// TIA Portal V20 export
// export: Created 2026-10-20T12:51:39.2775664Z, ExportSetting WithDefaults, DisplayName Totally Integrated Automation Portal, DisplayVersion V20 Update 6, DisplayName TIA Portal Openness, DisplayVersion V20 Update 6, DisplayName TIA Portal Version Control Interface, DisplayVersion V20 Update 6, DisplayName SINAMICS Startdrive Advanced, DisplayVersion V20 SP1, DisplayName SINAMICS Startdrive G130, G150, S120, S150, SINAMICS MV, G220, S200, S210, DisplayVersion V20 SP1, DisplayName SINAMICS Startdrive G110M, G120, G120C, G120D, G120P, G115D, DisplayVersion V20 SP1, DisplayName STEP 7 Professional, DisplayVersion V20 Update 6, DisplayName STEP 7 Safety, DisplayVersion V20 Update 2, DisplayName WinCC Basic/Comfort/Advanced, DisplayVersion V20 Update 6, DisplayName WinCC Unified, DisplayVersion V20 Update 6
FUNCTION "Bypass assignments_2" : Void   // FC36, F_LAD
{ S7_Optimized_Access := 'TRUE' }
VERSION : 0.1
// stored: AutoNumber true, IsIECCheckEnabled false, UDAEnableTagReadback false
BEGIN

REGION Network 1
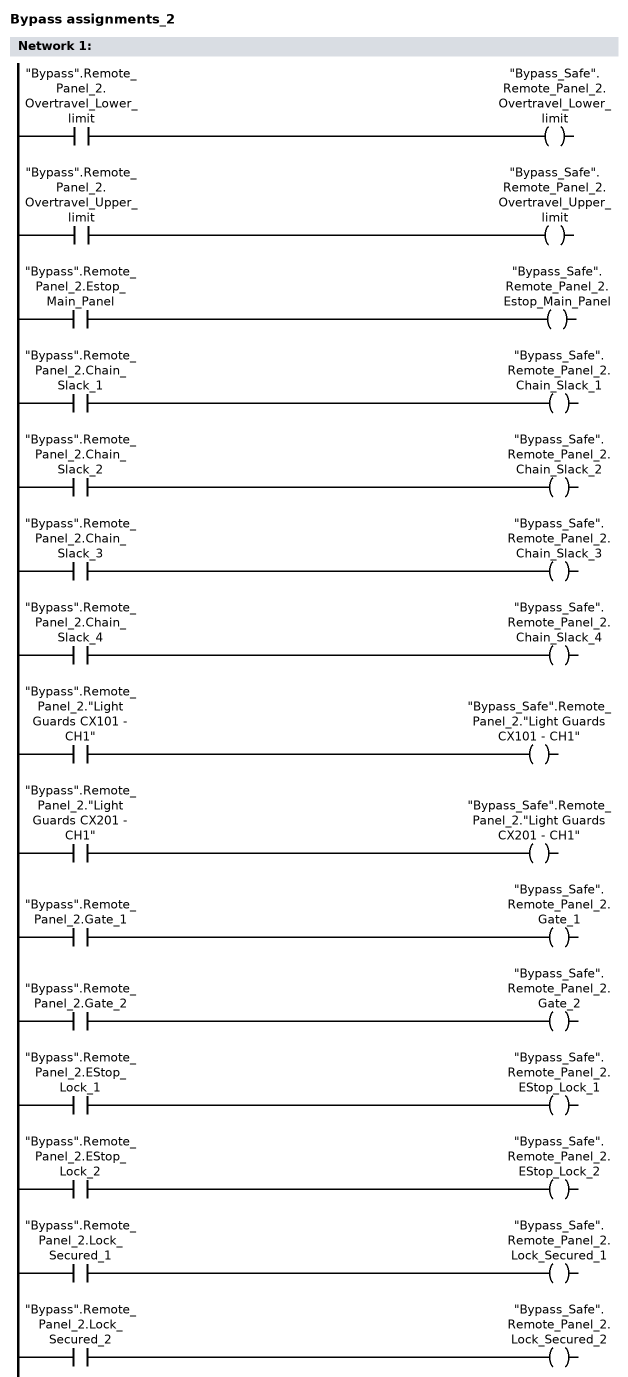
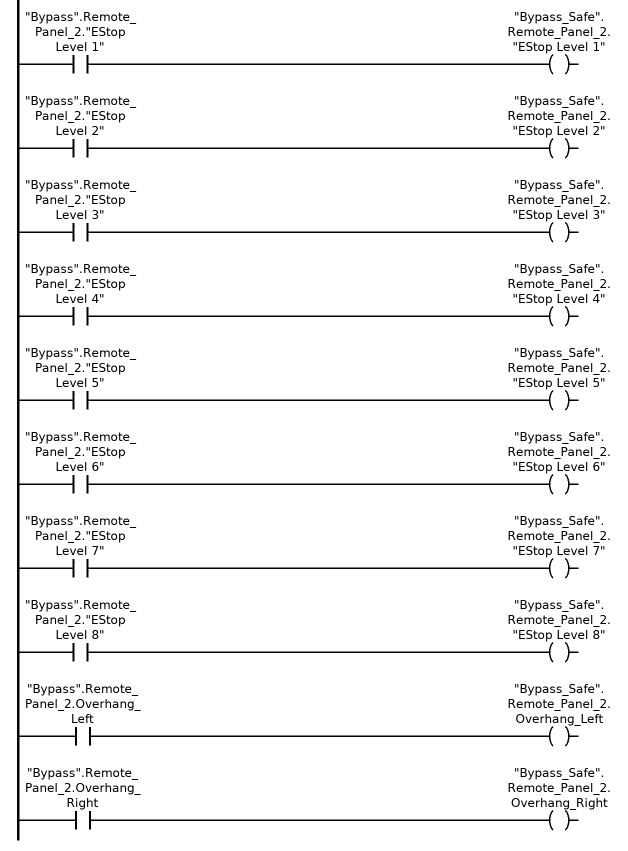
   RUNG wire#powerrail
      Contact( "Bypass".Remote_Panel_2.Overtravel_Lower_limit )
      Coil( "Bypass_Safe".Remote_Panel_2.Overtravel_Lower_limit )
   END_RUNG
   RUNG wire#powerrail
      Contact( "Bypass".Remote_Panel_2.Overtravel_Upper_limit )
      Coil( "Bypass_Safe".Remote_Panel_2.Overtravel_Upper_limit )
   END_RUNG
   RUNG wire#powerrail
      Contact( "Bypass".Remote_Panel_2.Estop_Main_Panel )
      Coil( "Bypass_Safe".Remote_Panel_2.Estop_Main_Panel )
   END_RUNG
   RUNG wire#powerrail
      Contact( "Bypass".Remote_Panel_2.Chain_Slack_1 )
      Coil( "Bypass_Safe".Remote_Panel_2.Chain_Slack_1 )
   END_RUNG
   RUNG wire#powerrail
      Contact( "Bypass".Remote_Panel_2.Chain_Slack_2 )
      Coil( "Bypass_Safe".Remote_Panel_2.Chain_Slack_2 )
   END_RUNG
   RUNG wire#powerrail
      Contact( "Bypass".Remote_Panel_2.Chain_Slack_3 )
      Coil( "Bypass_Safe".Remote_Panel_2.Chain_Slack_3 )
   END_RUNG
   RUNG wire#powerrail
      Contact( "Bypass".Remote_Panel_2.Chain_Slack_4 )
      Coil( "Bypass_Safe".Remote_Panel_2.Chain_Slack_4 )
   END_RUNG
   RUNG wire#powerrail
      Contact( "Bypass".Remote_Panel_2."Light Guards CX101 - CH1" )
      Coil( "Bypass_Safe".Remote_Panel_2."Light Guards CX101 - CH1" )
   END_RUNG
   RUNG wire#powerrail
      Contact( "Bypass".Remote_Panel_2."Light Guards CX201 - CH1" )
      Coil( "Bypass_Safe".Remote_Panel_2."Light Guards CX201 - CH1" )
   END_RUNG
   RUNG wire#powerrail
      Contact( "Bypass".Remote_Panel_2.Gate_1 )
      Coil( "Bypass_Safe".Remote_Panel_2.Gate_1 )
   END_RUNG
   RUNG wire#powerrail
      Contact( "Bypass".Remote_Panel_2.Gate_2 )
      Coil( "Bypass_Safe".Remote_Panel_2.Gate_2 )
   END_RUNG
   RUNG wire#powerrail
      Contact( "Bypass".Remote_Panel_2.EStop_Lock_1 )
      Coil( "Bypass_Safe".Remote_Panel_2.EStop_Lock_1 )
   END_RUNG
   RUNG wire#powerrail
      Contact( "Bypass".Remote_Panel_2.EStop_Lock_2 )
      Coil( "Bypass_Safe".Remote_Panel_2.EStop_Lock_2 )
   END_RUNG
   RUNG wire#powerrail
      Contact( "Bypass".Remote_Panel_2.Lock_Secured_1 )
      Coil( "Bypass_Safe".Remote_Panel_2.Lock_Secured_1 )
   END_RUNG
   RUNG wire#powerrail
      Contact( "Bypass".Remote_Panel_2.Lock_Secured_2 )
      Coil( "Bypass_Safe".Remote_Panel_2.Lock_Secured_2 )
   END_RUNG
   RUNG wire#powerrail
      Contact( "Bypass".Remote_Panel_2."EStop Level 1" )
      Coil( "Bypass_Safe".Remote_Panel_2."EStop Level 1" )
   END_RUNG
   RUNG wire#powerrail
      Contact( "Bypass".Remote_Panel_2."EStop Level 2" )
      Coil( "Bypass_Safe".Remote_Panel_2."EStop Level 2" )
   END_RUNG
   RUNG wire#powerrail
      Contact( "Bypass".Remote_Panel_2."EStop Level 3" )
      Coil( "Bypass_Safe".Remote_Panel_2."EStop Level 3" )
   END_RUNG
   RUNG wire#powerrail
      Contact( "Bypass".Remote_Panel_2."EStop Level 4" )
      Coil( "Bypass_Safe".Remote_Panel_2."EStop Level 4" )
   END_RUNG
   RUNG wire#powerrail
      Contact( "Bypass".Remote_Panel_2."EStop Level 5" )
      Coil( "Bypass_Safe".Remote_Panel_2."EStop Level 5" )
   END_RUNG
   RUNG wire#powerrail
      Contact( "Bypass".Remote_Panel_2."EStop Level 6" )
      Coil( "Bypass_Safe".Remote_Panel_2."EStop Level 6" )
   END_RUNG
   RUNG wire#powerrail
      Contact( "Bypass".Remote_Panel_2."EStop Level 7" )
      Coil( "Bypass_Safe".Remote_Panel_2."EStop Level 7" )
   END_RUNG
   RUNG wire#powerrail
      Contact( "Bypass".Remote_Panel_2."EStop Level 8" )
      Coil( "Bypass_Safe".Remote_Panel_2."EStop Level 8" )
   END_RUNG
   RUNG wire#powerrail
      Contact( "Bypass".Remote_Panel_2.Overhang_Left )
      Coil( "Bypass_Safe".Remote_Panel_2.Overhang_Left )
   END_RUNG
   RUNG wire#powerrail
      Contact( "Bypass".Remote_Panel_2.Overhang_Right )
      Coil( "Bypass_Safe".Remote_Panel_2.Overhang_Right )
   END_RUNG
   // the same network as SCL:
   "Bypass_Safe".Remote_Panel_2.Overtravel_Lower_limit := "Bypass".Remote_Panel_2.Overtravel_Lower_limit;
   "Bypass_Safe".Remote_Panel_2.Overtravel_Upper_limit := "Bypass".Remote_Panel_2.Overtravel_Upper_limit;
   "Bypass_Safe".Remote_Panel_2.Estop_Main_Panel := "Bypass".Remote_Panel_2.Estop_Main_Panel;
   "Bypass_Safe".Remote_Panel_2.Chain_Slack_1 := "Bypass".Remote_Panel_2.Chain_Slack_1;
   "Bypass_Safe".Remote_Panel_2.Chain_Slack_2 := "Bypass".Remote_Panel_2.Chain_Slack_2;
   "Bypass_Safe".Remote_Panel_2.Chain_Slack_3 := "Bypass".Remote_Panel_2.Chain_Slack_3;
   "Bypass_Safe".Remote_Panel_2.Chain_Slack_4 := "Bypass".Remote_Panel_2.Chain_Slack_4;
   "Bypass_Safe".Remote_Panel_2."Light Guards CX101 - CH1" := "Bypass".Remote_Panel_2."Light Guards CX101 - CH1";
   "Bypass_Safe".Remote_Panel_2."Light Guards CX201 - CH1" := "Bypass".Remote_Panel_2."Light Guards CX201 - CH1";
   "Bypass_Safe".Remote_Panel_2.Gate_1 := "Bypass".Remote_Panel_2.Gate_1;
   "Bypass_Safe".Remote_Panel_2.Gate_2 := "Bypass".Remote_Panel_2.Gate_2;
   "Bypass_Safe".Remote_Panel_2.EStop_Lock_1 := "Bypass".Remote_Panel_2.EStop_Lock_1;
   "Bypass_Safe".Remote_Panel_2.EStop_Lock_2 := "Bypass".Remote_Panel_2.EStop_Lock_2;
   "Bypass_Safe".Remote_Panel_2.Lock_Secured_1 := "Bypass".Remote_Panel_2.Lock_Secured_1;
   "Bypass_Safe".Remote_Panel_2.Lock_Secured_2 := "Bypass".Remote_Panel_2.Lock_Secured_2;
   "Bypass_Safe".Remote_Panel_2."EStop Level 1" := "Bypass".Remote_Panel_2."EStop Level 1";
   "Bypass_Safe".Remote_Panel_2."EStop Level 2" := "Bypass".Remote_Panel_2."EStop Level 2";
   "Bypass_Safe".Remote_Panel_2."EStop Level 3" := "Bypass".Remote_Panel_2."EStop Level 3";
   "Bypass_Safe".Remote_Panel_2."EStop Level 4" := "Bypass".Remote_Panel_2."EStop Level 4";
   "Bypass_Safe".Remote_Panel_2."EStop Level 5" := "Bypass".Remote_Panel_2."EStop Level 5";
   "Bypass_Safe".Remote_Panel_2."EStop Level 6" := "Bypass".Remote_Panel_2."EStop Level 6";
   "Bypass_Safe".Remote_Panel_2."EStop Level 7" := "Bypass".Remote_Panel_2."EStop Level 7";
   "Bypass_Safe".Remote_Panel_2."EStop Level 8" := "Bypass".Remote_Panel_2."EStop Level 8";
   "Bypass_Safe".Remote_Panel_2.Overhang_Left := "Bypass".Remote_Panel_2.Overhang_Left;
   "Bypass_Safe".Remote_Panel_2.Overhang_Right := "Bypass".Remote_Panel_2.Overhang_Right;
END_REGION
END_FUNCTION
